(* PLC project zarechnaya.project, CODESYS CODESYS V3.5 SP17 Patch 3 *)
(* stored: creationDateTime 2026-10-20T05:42:22.166614, modificationDateTime 1601-01-01T03:00:00 *)

(* F_Convert — пересчёт аналоговой уставки дозатора коагулянта (ST, FUNCTION). Поведение (по нему считает модель scenarios/reference/model_F_Convert.py): - результат функции — REAL_TO_INT(rIn): половина округляется от нуля (2.5 → 3, −2.5 → −3; проба M0); - iSum := iA + iB с переносом INT (32767 + 1 = −32768); - iQuot := iA / iB с отбрасыванием дробной части к нулю, при iB = 0 — 0 (делитель-переменная → C2S7-SEM-DIV0); - iMux := MUX(iSel, 10, 20, 30), iSel ∈ 0…2; - iLim := LIMIT(iMn, результат, iMx); при MN > MX результат — MX (проба M0: LIMIT(10, 5, 0) = 0). *)
FUNCTION F_Convert : INT
  VAR_INPUT
    rIn : REAL;
    iA : INT;
    iB : INT;
    iSel : INT;
    iMn : INT;
    iMx : INT;
  END_VAR
  VAR_OUTPUT
    iSum : INT;
    iQuot : INT;
    iMux : INT;
    iLim : INT;
  END_VAR

            F_Convert := REAL_TO_INT(rIn);
iSum := iA + iB;
IF iB <> 0 THEN
    iQuot := iA / iB;
ELSE
    iQuot := 0;
END_IF
iMux := MUX(iSel, 10, 20, 30);
iLim := LIMIT(iMn, F_Convert, iMx);

          
END_FUNCTION
